Staubli VAL3: progTemplate.dtx

public string sTRAJname
public num nType
public ifItem iIfItem
  [0]
    num nSigType[3]
    num nSigIndex[3]
    num nValue[3]
    bool bANDOR[2]
public switchItem sSwitchItem
  [0]
    num nSwitchValue
    string sIOValue
    bool bIOdisable
public forItem fForItem
  [0]
    num nLoopValue
    bool bIOdisable
    string sIOindex
    string sForTRAJ
